(* IEC 61131-3 sources: model-first-plc-agent-ai/results/T1-W-11, 2 files *)

(* ---- a1_code.st ---- *)
FUNCTION_BLOCK ConveyorRuntime
VAR_INPUT
    sensor_a : BOOL;
    sensor_b : BOOL;
END_VAR
VAR_OUTPUT
    conveyor : BOOL := FALSE;
END_VAR
VAR
    run_latch : RS;
END_VAR

(* The reset-dominant latch initializes FALSE, representing initial step x0.
   Its TRUE state represents step x1. *)
run_latch(
    S := sensor_a AND NOT sensor_b,
    R1 := sensor_b
);

conveyor := run_latch.Q1;

END_FUNCTION_BLOCK

PROGRAM Main
VAR
    SensorA AT %IX100.0 : BOOL;
    SensorB AT %IX100.1 : BOOL;
    Conveyor AT %QX100.0 : BOOL;
END_VAR
VAR
    runtime_logic : ConveyorRuntime;
END_VAR

(* Instance initialization establishes x0 before cyclic execution. *)
runtime_logic(
    sensor_a := SensorA,
    sensor_b := SensorB
);

Conveyor := runtime_logic.conveyor;

END_PROGRAM

(* ---- a2_code.st ---- *)
FUNCTION_BLOCK FB_ConveyorControl
VAR_INPUT
    sensor_a : BOOL;
    sensor_b : BOOL;
END_VAR
VAR_OUTPUT
    conveyor : BOOL;
END_VAR
VAR
    conveyor_latch : RS;
END_VAR

conveyor_latch(
    S := sensor_a AND NOT sensor_b,
    R1 := sensor_b
);
conveyor := conveyor_latch.Q1;

END_FUNCTION_BLOCK

PROGRAM Main
VAR
    sensor_a AT %IX100.0 : BOOL;
    sensor_b AT %IX100.1 : BOOL;
    conveyor AT %QX100.0 : BOOL;
END_VAR
VAR
    controller : FB_ConveyorControl;
END_VAR

controller(
    sensor_a := sensor_a,
    sensor_b := sensor_b
);
conveyor := controller.conveyor;

END_PROGRAM
